(*
SPDX-FileCopyrightText: c 2026 Oleksandr Tiutyk <trofimich@gmail.com>
SPDX-License-Identifier: MIT
License: https://opensource.org/license/mit
*)

(*!
<summary>Checks the current LIFO top and length after each push.</summary>
<description>
Borrows a group-owned stack reserved for this case. Use from one task at a stable address.
Teardown clears the stack and test-owned resources before publication.
</description>
*)

{attribute 'no_assign'}
{attribute 'no_explicit_call' := 'do not call this function block directly'}
FUNCTION_BLOCK StackPushAndPeekTest EXTENDS TOF_Testing.SingleCycleTest
VAR_STAT
	{attribute 'hide'}
	_ClassName : STRING := __POUNAME();
END_VAR
VAR
	_Stack : TOF_Collections.IStack;
END_VAR

(*!
<summary>Clears the fixture before the runner publishes the result.</summary>
<description>
Also runs after an unexpected exception interrupts the case.
</description>
*)
METHOD PROTECTED AfterTest
_Stack.Clear();
END_METHOD

//! <summary>Borrows the concrete class name. Callers must not modify it.</summary>
{attribute 'monitoring' := 'call'}
PROPERTY ClassName : REFERENCE TO STRING
GET
ClassName REF= _ClassName;
END_GET
END_PROPERTY

(*!
<summary>Checks the current LIFO top and length after each push.</summary>
*)
METHOD PROTECTED ExecuteTest
VAR
	values : ARRAY [1..4] OF INT := [11, 22, 33, 44];
END_VAR
_Stack.PushCopy(value := values[1]);

Assert.ThatInt(
	actual := _Stack.Peek().AsInt(),
	message := "Push 1 must establish the new top"
).ToBe(expected := values[1]);

Assert.ThatDInt(
	actual := _Stack.Length,
	message := "Peeking after push 1 must preserve length"
).ToBe(expected := DINT#1);

_Stack.PushCopy(value := values[2]);

Assert.ThatInt(
	actual := _Stack.Peek().AsInt(),
	message := "Push 2 must establish the new top"
).ToBe(expected := values[2]);

Assert.ThatDInt(
	actual := _Stack.Length,
	message := "Peeking after push 2 must preserve length"
).ToBe(expected := DINT#2);

_Stack.PushCopy(value := values[3]);

Assert.ThatInt(
	actual := _Stack.Peek().AsInt(),
	message := "Push 3 must establish the new top"
).ToBe(expected := values[3]);

Assert.ThatDInt(
	actual := _Stack.Length,
	message := "Peeking after push 3 must preserve length"
).ToBe(expected := DINT#3);
END_METHOD

(*!
<summary>Binds the stack fixture for this case.</summary>
<description>
Stores a borrowed interface without invoking the fixture. The owning group keeps it alive and
reserves it for this case. TestElement initializes the name and parent.
</description>
<param name="name">Display name of this case.</param>
<param name="parent">Group that owns this case.</param>
<param name="stack">Required live stack reserved for this case.</param>
*)
METHOD FB_init : BOOL
VAR_INPUT
	bInitRetains: BOOL; // TRUE: the retain variables are initialized (reset warm / reset cold)
	bInCopyCode: BOOL; // TRUE: the instance will be copied to the copy code afterward (online change)
	name : WSTRING;
	parent : TOF_Testing.ITestElement;
	stack : TOF_Collections.IStack;
END_VAR
_Stack := stack;
FB_init := TRUE;
END_METHOD

//! <summary>Borrows the compiler-initialized namespace name. Callers must not modify it.</summary>
{attribute 'monitoring' := 'call'}
PROPERTY NamespaceName : REFERENCE TO STRING
GET
NamespaceName REF= CurrentNamespace.Name;
END_GET
END_PROPERTY

//! <summary>Reports the concrete instance size in bytes.</summary>
{attribute 'monitoring' := 'call'}
PROPERTY SelfSize : ULINT
GET
SelfSize := XSIZEOF(THIS^);
END_GET
END_PROPERTY

END_FUNCTION_BLOCK

(* stored: Version 1.1.0.1, ProductVersion 3.1.4026.21
   POU StackPushAndPeekTest: Id {1e0f0d81-b6ea-4997-b2d6-74d7a036653a}, SpecialFunc None
   Method AfterTest: Id {4e72989c-514a-4e22-8217-0c61fb5d6269}
   Property ClassName: Id {d6843c90-ec27-41dd-ac88-4813e63c8e37}
   Get Get: Id {5bc9100c-800b-4bcb-9d59-97faa9c41aee}
   Method ExecuteTest: Id {1f43e591-99f6-449f-bd73-90cdf35f4916}
   Method FB_init: Id {883f9d39-5611-4c97-9a4e-52c630b8ee33}
   Property NamespaceName: Id {7b6fc482-d81e-4b1d-b1a2-171c65516c36}
   Get Get: Id {2b2c3a10-b909-47c3-b2a5-3ffd34654e08}
   Property SelfSize: Id {e137269f-756a-42e8-88e3-b565e12e83de}
   Get Get: Id {b24afb9e-2504-4a59-975a-936af3decb5d} *)
